(* IEC 61131-3 sources: 308sjk/scenegen/out/plotter_cell_draw, 1 file *)

(* ---- st_io_declaration.st ---- *)
VAR_GLOBAL
    x_fb AT %QW0 : INT;   (* 输入反馈：工程量定点 int16，换算归桥 *)
    y_fb AT %QW1 : INT;   (* 输入反馈：工程量定点 int16，换算归桥 *)
    z_fb AT %QW2 : INT;   (* 输入反馈：工程量定点 int16，换算归桥 *)
END_VAR
